(* IEC 61131-3 sources: kns-port-domestic/targets/astra/src/DUTs/Log, 8 files *)

(* ---- E_EventKind.dut.st ---- *)
// Назначение: вид записи журнала (ST_EventRecord.eKind): событие тревоги PL.FB_Alarm или событие станции.
// Автор:      kr0nsch
// Версия:     0.1.0
// Документ:   docs/DESIGN.md, раздел 3.2
{attribute 'qualified_only'}
{attribute 'strict'}
TYPE E_EventKind :
(
    Alarm   := 1,   // переход тревоги (PL.I_AlarmSink.OnAlarmEvent)
    Station := 2    // событие станции (I_StationEventSink.LogEvent), номер 101000 + код
) INT;
END_TYPE

(* ---- E_LogExportState.dut.st ---- *)
// Назначение: состояние выгрузки журнала в CSV (GVL_Log.eExportState, stStationSts.eLogExport).
// Автор:      kr0nsch
// Версия:     0.1.0
// Документ:   docs/DESIGN.md, раздел 3.2
{attribute 'qualified_only'}
{attribute 'strict'}
TYPE E_LogExportState :
(
    Idle     := 0,   // выгрузки не было
    Snapshot := 1,   // снимок кольца сделан, ждёт SlowTask
    Writing  := 2,   // SlowTask пишет файл
    Done     := 3,   // файл записан
    Error    := 4    // ошибка CAA File
) INT;
END_TYPE

(* ---- E_StationEvent.dut.st ---- *)
// Назначение: события станции в журнале (04 §16): номер записи = STN_EVENT_ID_BASE + код.
//             Без strict: значение кода пишется в журнал числом (DESIGN, раздел 3.2).
// Автор:      kr0nsch
// Версия:     0.1.0
// Документ:   docs/DESIGN.md, раздел 3.2
{attribute 'qualified_only'}
TYPE E_StationEvent :
(
    StationAuto       := 1,    // режим станции «Автомат»
    StationManual     := 2,    // режим станции «Ручной»
    MethodStepped     := 3,    // способ: ступенчатое
    MethodLevelPid    := 4,    // способ: ПИД уровня
    LeadChanged       := 5,    // смена ведущего (номер насоса)
    AtsPumpIn         := 6,    // АВР: введён насос (номер насоса)
    ContRunHandover   := 7,    // передача роли по ограничению непрерывной работы (номер нового насоса)
    PowerLost         := 8,    // пропадание напряжения
    RestartBegin      := 9,    // начало последовательного пуска
    RestartDone       := 10,   // последовательный пуск завершён (число пущенных)
    FloatMasked       := 11,   // поплавок исключён (102 или 103)
    FloatUnmasked     := 12,   // поплавок возвращён (102 или 103)
    FloatModeOn       := 13,   // переход на управление по поплавкам
    FloatModeOff      := 14,   // возврат к управлению по LT101
    PlcStart          := 15,   // старт приложения ПЛК
    ResetAll          := 16,   // общий сброс (1 — кнопка, 2 — HMI)
    CfgChanged        := 17,   // изменение уставки станции (номер параметра)
    DeviceModeChanged := 18,   // смена режима устройства (dev_no * 10 + режим)
    LogExported       := 19,   // журнал выгружен (строк)
    LogExportFailed   := 20,   // ошибка выгрузки (код ошибки CAA File)
    SimFaultChanged   := 21,   // изменена инъекция отказа (номер поля)
    AckAll            := 22,   // квитировать все
    Silence           := 23    // звук отключён (1 — кнопка, 2 — HMI)
) UINT;
END_TYPE

(* ---- ST_AlarmView.dut.st ---- *)
// Назначение: список тревог не в Normal (GVL_Log.stAlarmView): неквитированные выше, затем активные по
//             приоритету, затем подавленные и отложенные, внутри группы — новые выше.
// Автор:      kr0nsch
// Версия:     0.1.0
// Документ:   docs/DESIGN.md, раздел 3.2
{attribute 'qualified_only'}
TYPE ST_AlarmView :
STRUCT
    uiCount       : UINT;           // строк в astRow
    uiActiveTotal : UINT;           // настоящее число тревог не в Normal (может быть больше ALM_VIEW_ROWS)
    udiRevision   : UDINT;          // +1 при каждом пересчёте
    astRow        : ARRAY[1..GVL_Const.ALM_VIEW_ROWS] OF ST_AlarmViewRow;
END_STRUCT
END_TYPE

(* ---- ST_AlarmViewRow.dut.st ---- *)
// Назначение: строка списка тревог не в Normal (баннер, экран «Тревоги», сценарии ПМИ).
// Автор:      kr0nsch
// Версия:     0.1.0
// Документ:   docs/DESIGN.md, раздел 3.2
{attribute 'qualified_only'}
TYPE ST_AlarmViewRow :
STRUCT
    udiId          : UDINT;
    ePriority      : PL.E_AlarmPriority;
    eState         : PL.E_AlarmState;
    uiSource       : UINT;          // индекс источника в FB_AlarmSummary (устройства — индекс GVL_DeviceList)
    uiSlot         : UINT;
    uliSinceUtc_ms : ULINT;         // время последнего перехода, замеченного сводкой
END_STRUCT
END_TYPE

(* ---- ST_EventFeed.dut.st ---- *)
// Назначение: курсор журнала для внешних клиентов (GVL_Log.stEventFeed: сценарии ПМИ, SCADA) — записи от
//             старой к новой начиная с номера udiFromSeq, отдельно от страницы HMI. Клиент читает строки,
//             пишет udiFromSeq := номер последней прочитанной + 1 и повторяет; udiFromSeq < udiSeqFirst —
//             записи между опросами затёрты (пропуск номеров).
// Автор:      kr0nsch
// Версия:     0.1.0
// Документ:   docs/DESIGN.md, разделы 3.2, 14.3
{attribute 'qualified_only'}
TYPE ST_EventFeed :
STRUCT
    udiFromSeq  : UDINT;            // пишет клиент: первый нужный номер
    udiSeqFirst : UDINT;            // самая старая запись в кольце (пустой журнал — udiSeqLast + 1)
    udiSeqLast  : UDINT;            // самая новая запись (0 — записей ещё не было)
    uiCount     : UINT;             // строк в astRow
    wReserve    : WORD;
    astRow      : ARRAY[1..GVL_Const.LOG_FEED_ROWS] OF ST_EventRecord;   // строки после uiCount — нули
END_STRUCT
END_TYPE

(* ---- ST_EventRecord.dut.st ---- *)
// Назначение: запись журнала событий FB_EventLog (кольцо LOG_CAPACITY записей). 40 байт: 32-битные поля
//             на смещениях, кратных 4, ULINT и LREAL — кратных 8 (тест EventRecordSizeIs40).
// Автор:      kr0nsch
// Версия:     0.1.0
// Документ:   docs/DESIGN.md, раздел 3.2
{attribute 'qualified_only'}
TYPE ST_EventRecord :
STRUCT
    udiSeq    : UDINT;                  // сквозной номер с запуска приложения, с 1
    eKind     : E_EventKind;
    ePriority : PL.E_AlarmPriority;     // события станции — None
    udiId     : UDINT;                  // номер тревоги или 101000 + код события
    eOldState : PL.E_AlarmState;        // события станции — Normal
    eNewState : PL.E_AlarmState;
    eReason   : PL.E_AlarmEventReason;  // события станции — None
    wReserve  : WORD;                   // выравнивание: дальше 32- и 64-битные поля
    rValue    : REAL;                   // значение процесса или аргумент события
    uliUtc_ms : ULINT;                  // UTC, мс от 1970 (SysTimeRtcHighResGet); 0 — часы недоступны
    lrMono_s  : LREAL;                  // время процесса, с (I_TimeSource журнала = GVL_Time.fbClockMain)
END_STRUCT
END_TYPE

(* ---- ST_EventView.dut.st ---- *)
// Назначение: страница журнала для HMI (GVL_Log.stEventView): новые записи сверху, uiPage пишет HMI.
// Автор:      kr0nsch
// Версия:     0.1.0
// Документ:   docs/DESIGN.md, раздел 3.2
{attribute 'qualified_only'}
TYPE ST_EventView :
STRUCT
    uiPage      : UINT;             // пишет HMI: 0 — новые; больше последней — последняя страница
    uiPageCount : UINT;             // страниц (не меньше 1)
    uiCount     : UINT;             // записей в журнале
    wReserve    : WORD;
    astRow      : ARRAY[1..GVL_Const.LOG_VIEW_ROWS] OF ST_EventRecord;   // пустые строки — udiSeq = 0
END_STRUCT
END_TYPE
